(* IEC 61131-3 sources: plc-sbom-builder/samples/maschine-xy/programm/Verpackung, 1 file *)

(* ---- PLC_PRG.st ---- *)
PROGRAM PLC_PRG
VAR
    bStart : BOOL;
    nTakt : INT;
END_VAR

IF bStart THEN
    nTakt := nTakt + 1;
END_IF
